{attribute 'reflection'}
FUNCTION_BLOCK FB_GaugeBase
VAR
    //Logging
    fbLogger : FB_LogMessage := (eSubsystem:=E_SubSystem.VACUUM);
    ePrevState : E_PressureState;
    tErrorPresent : R_TRIG;
    tAction : R_TRIG; // Primary action of this device (OPN_DO, etc.)
    tOverrideActivated : R_TRIG;
     tState : R_TRIG;
    {attribute 'instance-path'}
    {attribute 'noinit'}
    sPath: STRING;
    // For Persistent Data
    bRestorePersistentData	:	BOOL:=TRUE;
    stateTimer:TON;
    fbGetCurTaskIdx  : GETCURTASKINDEX;
    fbWritePersistentData           : WritePersistentData;
    tRecover: TON;
END_VAR
VAR PERSISTENT
    rVAC_SP	:	REAL;
    rPRO_SP	:	REAL;
    rHYS_PR: REAL;
END_VAR

END_FUNCTION_BLOCK

(* stored: Version 1.1.0.1
   POU FB_GaugeBase: Id {7a1f28cc-0783-4ebe-9457-6569085eece6}, SpecialFunc None *)
